(* PLC project Storage_Main, Beckhoff Automation GmbH TwinCAT PLC Control 3.5.13.21 *)
(* stored: creationDateTime 2026-11-24T10:16:09.8423359, modificationDateTime 2026-11-24T10:16:09.8423359 *)

PROGRAM SFC_T1
// =====================================================================
// SFC_T1 (Sequential Function Chart)
// Homing and the automatic sequence (GRAFCET E70 .. S70).
// Called from MAIN every cycle. All variables are in MAIN (MAIN.xxx).
// Every step has one ST action (<step>_Active) that runs while the step is active.
// The motors are switched off in MAIN before this chart is called, so a step
// only has to switch ON what it needs.
// =====================================================================
VAR_INPUT
    SFCReset : BOOL;            // SFC flag: TRUE = chart back to the initial step S0 (STOP / homing timeout)
END_VAR
VAR
END_VAR

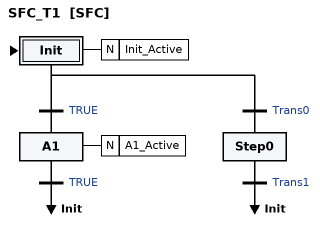
INITIAL_STEP Init:
  Init_Active(N);
END_STEP
TRANSITION FROM Init TO A1
  := TRUE;
END_TRANSITION
TRANSITION FROM Init TO Step0
  := Trans0;
END_TRANSITION
STEP Step0:
END_STEP
TRANSITION FROM Step0 TO Init
  := Trans1;
END_TRANSITION
STEP A1:
  A1_Active(N);
END_STEP
TRANSITION FROM A1 TO Init
  := TRUE;
END_TRANSITION

ACTION Init_Active:
                MAIN.nStep := MAIN.nStep;
              
END_ACTION

ACTION A1_Active:
                MAIN.nStep := MAIN.nStep;
              
END_ACTION
END_PROGRAM
